(* Logix 5000 project; controller TFF vendor 1 type 14 code 107 rev 33.11; software revision 33.04; part 30 of 38 *)
(* tags used below, declared in another part *)
   Index : DINT;   // Index
   AA008 : ALIAS FOR DigitalPoint[18];
   AI101 : ALIAS FOR AnalogPoint[16];
   AI101_SIG : ALIAS FOR DigitalPoint[106];
   AI104 : ALIAS FOR AnalogPoint[17];
   AI104_SIG : ALIAS FOR DigitalPoint[107];
   AI201B : ALIAS FOR AnalogPoint[0];
   AI201B_SIG : ALIAS FOR DigitalPoint[109];
   AI202 : ALIAS FOR AnalogPoint[9];
   AI202_SIG : ALIAS FOR DigitalPoint[105];
   ARC_AI101 : ARC_pH;
   ARC_AI202 : ARC_pH;
   DF24VDC : ALIAS FOR DigitalPoint[4];
   DF24VDCPC : ALIAS FOR DigitalPoint[25];
   DF3PHP003 : ALIAS FOR DigitalPoint[27];
   DigitalInput : BOOL[256];   // Digital Input Array these bits are copied from Input cards.
   DigitalPoint : DigitalPoint[150];   // Digital Point Array
   ES001 : ALIAS FOR DigitalPoint[2];
   FI101 : ALIAS FOR AnalogPoint[19];
   FI101_SIG : ALIAS FOR DigitalPoint[110];
   MIX101 : ALIAS FOR AnalogPoint[14];
   MIX101_SIG : ALIAS FOR DigitalPoint[104];
   MIX101DF : ALIAS FOR DigitalPoint[28];
   Mixer : Mixer;   // Mixer config. structure
   Options : Options;   // Options List
   PCV101 : ALIAS FOR AnalogPoint[3];
   PCV101_SIG : ALIAS FOR DigitalPoint[102];
   PCV201 : ALIAS FOR AnalogPoint[4];
   PCV201_SIG : ALIAS FOR DigitalPoint[103];
   PI101 : ALIAS FOR AnalogPoint[6];
   PI101_SIG : ALIAS FOR DigitalPoint[98];
   PI201 : ALIAS FOR AnalogPoint[7];
   PI201_SIG : ALIAS FOR DigitalPoint[99];
   PI401 : ALIAS FOR AnalogPoint[8];
   PI401_SIG : ALIAS FOR DigitalPoint[100];
   PSH001 : ALIAS FOR DigitalPoint[21];
   PSH401 : ALIAS FOR DigitalPoint[22];
   Rack_Murr_Node0_Smart : IO_Station;   // Status of Node 0 Smart
   Rack_Murr_Node1_TFF20 : IO_Station;   // Status of Node 1 TFF20
   Rack_Murr_Node1_TFF40 : IO_Station;   // Status of Node 1 TFF40
   Rack_Murr_Node1_TFF80 : IO_Station;   // Status of Node 1 TFF80
   RSBUZZ : ALIAS FOR DigitalPoint[3];
   SIC001DF : ALIAS FOR DigitalPoint[16];
   SIC002DF : ALIAS FOR DigitalPoint[17];
   SIC003DF : ALIAS FOR DigitalPoint[29];
   TCU101 : ALIAS FOR AnalogPoint[18];
   TCU101_SIG : ALIAS FOR DigitalPoint[108];
   TCU101DF : ALIAS FOR DigitalPoint[30];
   ThisSystem : SystemType;
   TI101 : ALIAS FOR AnalogPoint[13];
   TI101_SIG : ALIAS FOR DigitalPoint[101];
   TI201 : ALIAS FOR AnalogPoint[22];
   TI201_SIG : ALIAS FOR DigitalPoint[111];
   ValveSwInput : BOOL[64];   // Valve digital input
   XS011 : ALIAS FOR DigitalPoint[14];
   XS012 : ALIAS FOR DigitalPoint[15];
   XV003 : ALIAS FOR Valve[2];
   XV004 : ALIAS FOR Valve[3];
   XV005 : ALIAS FOR Valve[4];
   XV006 : ALIAS FOR Valve[5];
   XV007 : ALIAS FOR Valve[6];
   ZS001 : ALIAS FOR DigitalPoint[6];
   ZS002 : ALIAS FOR DigitalPoint[7];
   ZS003 : ALIAS FOR DigitalPoint[8];
   ZS004 : ALIAS FOR DigitalPoint[9];
   ZS005 : ALIAS FOR DigitalPoint[10];
   ZS008 : ALIAS FOR DigitalPoint[5];
(* Process, continued *)

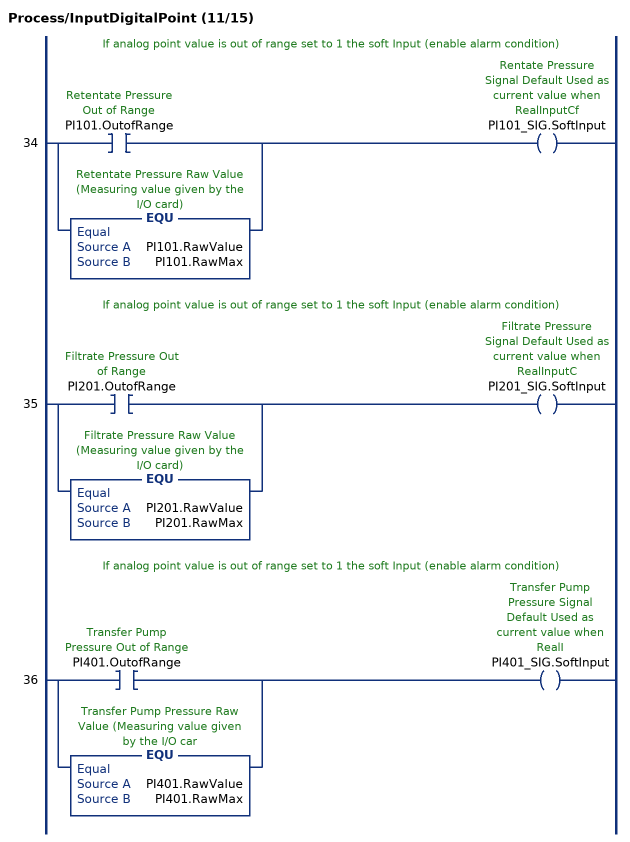
   [picture p330: Process/InputDigitalPoint rungs 34-36]
   // If analog point value is out of range set to 1 the soft Input (enable alarm condition)
   34: [XIC(PI101.OutofRange) ,EQU(PI101.RawValue,PI101.RawMax) ]OTE(PI101_SIG.SoftInput);
   // If analog point value is out of range set to 1 the soft Input (enable alarm condition)
   35: [XIC(PI201.OutofRange) ,EQU(PI201.RawValue,PI201.RawMax) ]OTE(PI201_SIG.SoftInput);
   // If analog point value is out of range set to 1 the soft Input (enable alarm condition)
   36: [XIC(PI401.OutofRange) ,EQU(PI401.RawValue,PI401.RawMax) ]OTE(PI401_SIG.SoftInput);
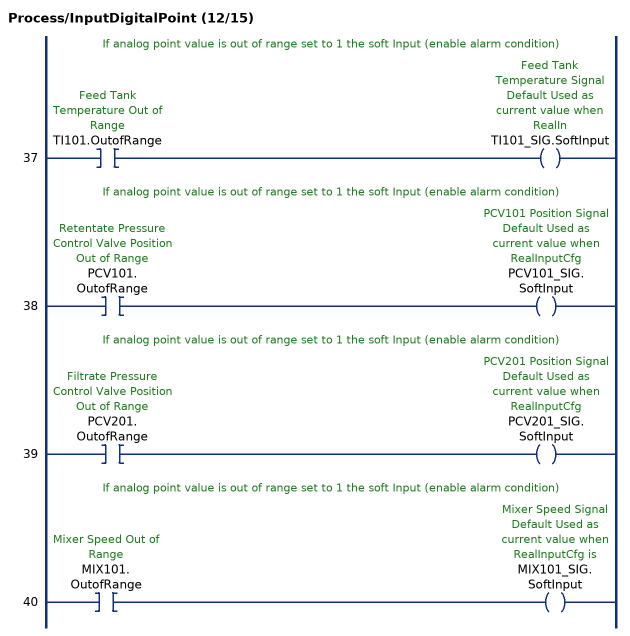
   // If analog point value is out of range set to 1 the soft Input (enable alarm condition)
   37: XIC(TI101.OutofRange)OTE(TI101_SIG.SoftInput);
   // If analog point value is out of range set to 1 the soft Input (enable alarm condition)
   38: XIC(PCV101.OutofRange)OTE(PCV101_SIG.SoftInput);
   // If analog point value is out of range set to 1 the soft Input (enable alarm condition)
   39: XIC(PCV201.OutofRange)OTE(PCV201_SIG.SoftInput);
   // If analog point value is out of range set to 1 the soft Input (enable alarm condition)
   40: XIC(MIX101.OutofRange)OTE(MIX101_SIG.SoftInput);
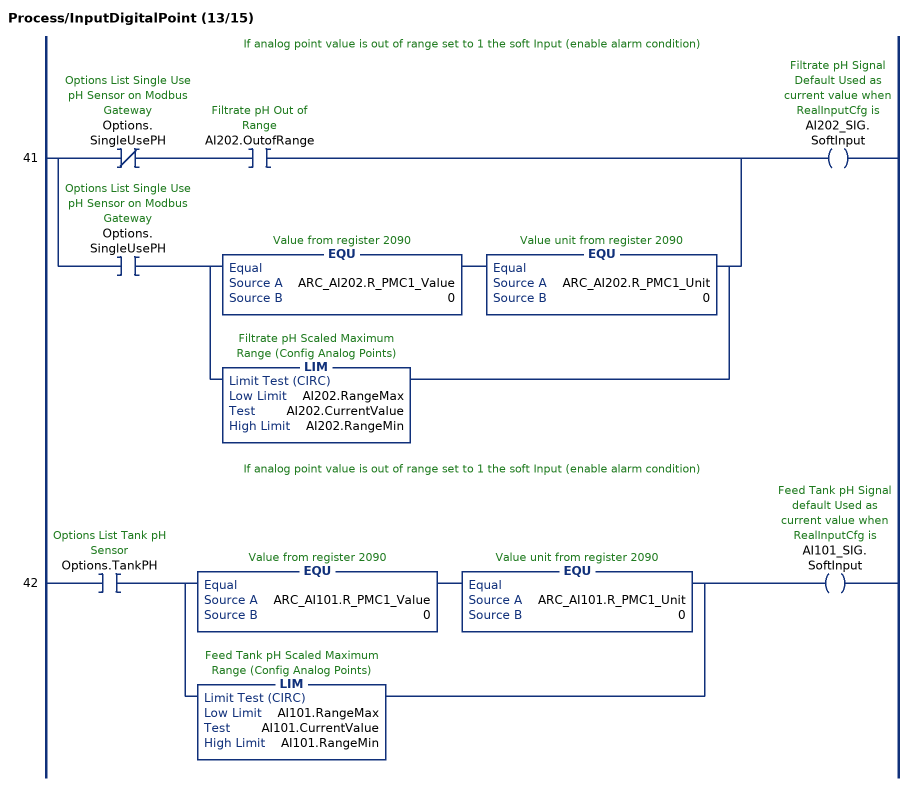
   // If analog point value is out of range set to 1 the soft Input (enable alarm condition)
   41: [XIO(Options.SingleUsePH) XIC(AI202.OutofRange) ,XIC(Options.SingleUsePH) [EQU(ARC_AI202.R_PMC1_Value,0) EQU(ARC_AI202.R_PMC1_Unit,0) ,LIM(AI202.RangeMax,AI202.CurrentValue,AI202.RangeMin) ] ]OTE(AI202_SIG.SoftInput);
   // If analog point value is out of range set to 1 the soft Input (enable alarm condition)
   42: XIC(Options.TankPH)[EQU(ARC_AI101.R_PMC1_Value,0) EQU(ARC_AI101.R_PMC1_Unit,0) ,LIM(AI101.RangeMax,AI101.CurrentValue,AI101.RangeMin) ]OTE(AI101_SIG.SoftInput);
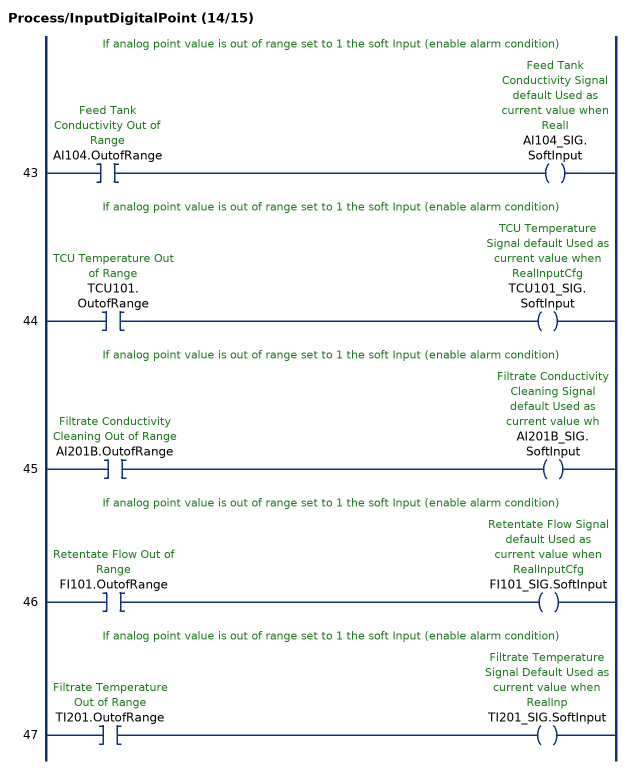
   // If analog point value is out of range set to 1 the soft Input (enable alarm condition)
   43: XIC(AI104.OutofRange)OTE(AI104_SIG.SoftInput);
   // If analog point value is out of range set to 1 the soft Input (enable alarm condition)
   44: XIC(TCU101.OutofRange)OTE(TCU101_SIG.SoftInput);
   // If analog point value is out of range set to 1 the soft Input (enable alarm condition)
   45: XIC(AI201B.OutofRange)OTE(AI201B_SIG.SoftInput);
   // If analog point value is out of range set to 1 the soft Input (enable alarm condition)
   46: XIC(FI101.OutofRange)OTE(FI101_SIG.SoftInput);
   // If analog point value is out of range set to 1 the soft Input (enable alarm condition)
   47: XIC(TI201.OutofRange)OTE(TI201_SIG.SoftInput);
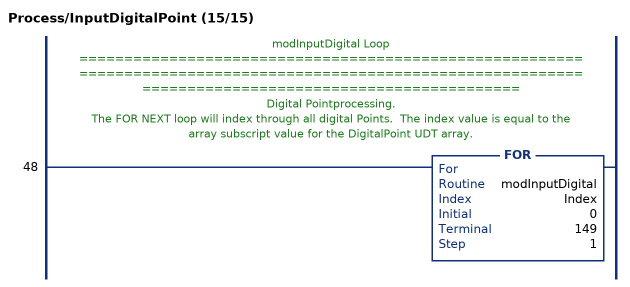
   // modInputDigital Loop
   // ==========================================================================================================================================================
   // Digital Pointprocessing.
   // The FOR NEXT loop will index through all digital Points.  The index value is equal to the array subscript value for the DigitalPoint UDT array.
   48: FOR(modInputDigital,Index,0,149,1);
END_ROUTINE

ROUTINE InputDigitalRaw   (* ladder *)
// Digital Input Routine
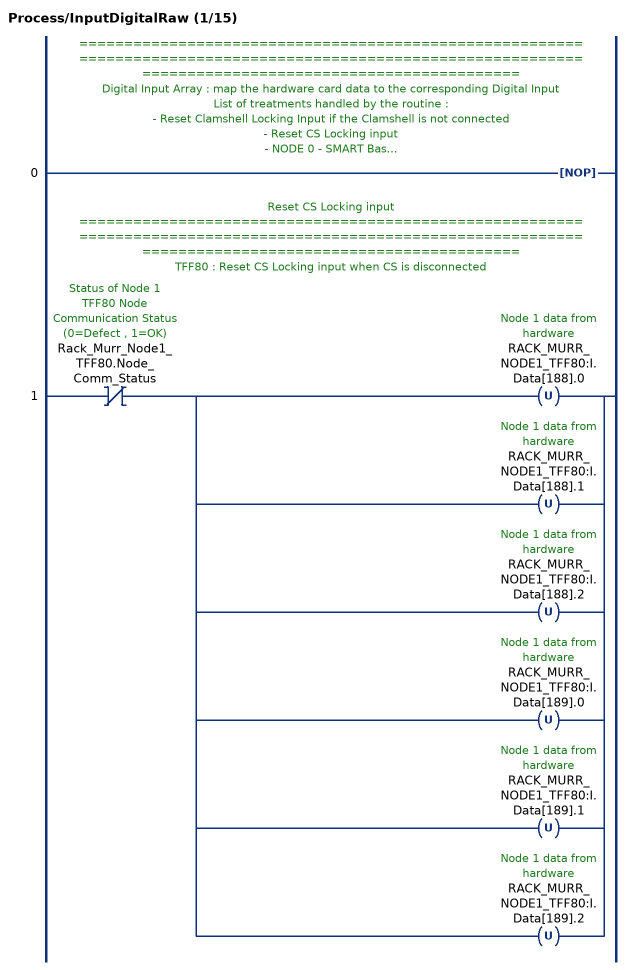
   // ==========================================================================================================================================================
   //                                                                                             Digital Input Array : map the hardware card data to the corresponding Digital Input
   //                                                     List of treatments handled by the routine :
   //                                                    - Reset Clamshell Locking Input if the Clamshell is not connected
   //                                                    - Reset CS Locking input
   //                                                    - NODE 0 - SMART Base
   //                                                         - NODE 1 - TFF80 Clamshell
   //                                                         - NODE 1 - TFF40 Clamshell
   //                                                         - NODE 1 - TFF20 Clamshell
   //                                                     -----------------------------------------------------------------------------------------------------------------------------------------------------
   //                                                     History
   // 		2019-DEC-24 - Merck - Q. Spindler - Initial version for Candidate Release 1.00.00.00.a
   // 		2020-APR-15 - Merck - Q. Spindler - Modifications for Candidate Release 1.00.00.00.b
   // - Add XS003, XS004, XS005, XS006, and XS007
   // ==========================================================================================================================================================
   0: NOP();
   // Reset CS Locking input
   // ==========================================================================================================================================================
   // TFF80 : Reset CS Locking input when CS is disconnected
   1: XIO(Rack_Murr_Node1_TFF80.Node_Comm_Status)[OTU(RACK_MURR_NODE1_TFF80:I.Data[188].0) ,OTU(RACK_MURR_NODE1_TFF80:I.Data[188].1) ,OTU(RACK_MURR_NODE1_TFF80:I.Data[188].2) ,OTU(RACK_MURR_NODE1_TFF80:I.Data[189].0) ,OTU(RACK_MURR_NODE1_TFF80:I.Data[189].1) ,OTU(RACK_MURR_NODE1_TFF80:I.Data[189].2) ];
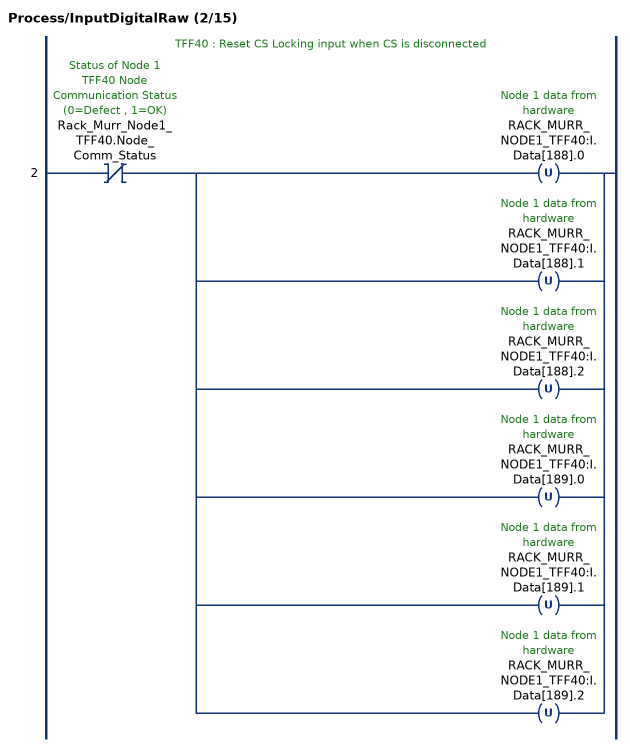
   // TFF40 : Reset CS Locking input when CS is disconnected
   2: XIO(Rack_Murr_Node1_TFF40.Node_Comm_Status)[OTU(RACK_MURR_NODE1_TFF40:I.Data[188].0) ,OTU(RACK_MURR_NODE1_TFF40:I.Data[188].1) ,OTU(RACK_MURR_NODE1_TFF40:I.Data[188].2) ,OTU(RACK_MURR_NODE1_TFF40:I.Data[189].0) ,OTU(RACK_MURR_NODE1_TFF40:I.Data[189].1) ,OTU(RACK_MURR_NODE1_TFF40:I.Data[189].2) ];
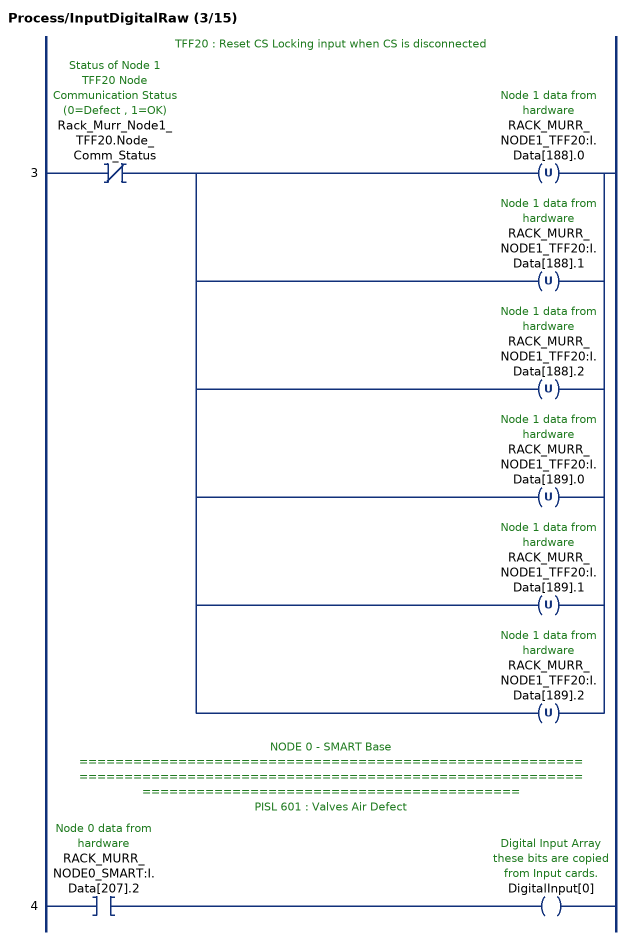
   // TFF20 : Reset CS Locking input when CS is disconnected
   3: XIO(Rack_Murr_Node1_TFF20.Node_Comm_Status)[OTU(RACK_MURR_NODE1_TFF20:I.Data[188].0) ,OTU(RACK_MURR_NODE1_TFF20:I.Data[188].1) ,OTU(RACK_MURR_NODE1_TFF20:I.Data[188].2) ,OTU(RACK_MURR_NODE1_TFF20:I.Data[189].0) ,OTU(RACK_MURR_NODE1_TFF20:I.Data[189].1) ,OTU(RACK_MURR_NODE1_TFF20:I.Data[189].2) ];
   // NODE 0 - SMART Base
   // ==========================================================================================================================================================
   // PISL 601 : Valves Air Defect
   4: XIC(RACK_MURR_NODE0_SMART:I.Data[207].2)OTE(DigitalInput[0]);
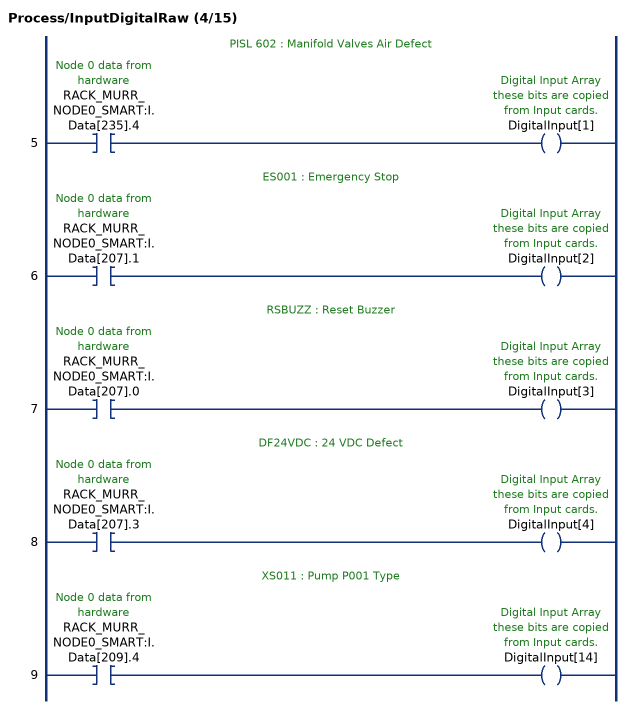
   // PISL 602 : Manifold Valves Air Defect
   5: XIC(RACK_MURR_NODE0_SMART:I.Data[235].4)OTE(DigitalInput[1]);
   // ES001 : Emergency Stop
   6: XIC(RACK_MURR_NODE0_SMART:I.Data[207].1)OTE(DigitalInput[2]);
   // RSBUZZ : Reset Buzzer
   7: XIC(RACK_MURR_NODE0_SMART:I.Data[207].0)OTE(DigitalInput[3]);
   // DF24VDC : 24 VDC Defect
   8: XIC(RACK_MURR_NODE0_SMART:I.Data[207].3)OTE(DigitalInput[4]);
   // XS011 : Pump P001 Type
   9: XIC(RACK_MURR_NODE0_SMART:I.Data[209].4)OTE(DigitalInput[14]);
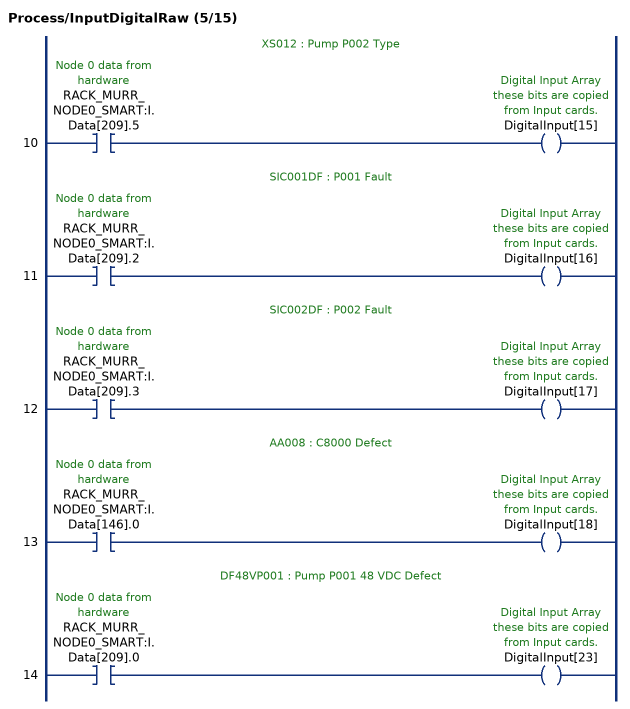
   // XS012 : Pump P002 Type
   10: XIC(RACK_MURR_NODE0_SMART:I.Data[209].5)OTE(DigitalInput[15]);
   // SIC001DF : P001 Fault
   11: XIC(RACK_MURR_NODE0_SMART:I.Data[209].2)OTE(DigitalInput[16]);
   // SIC002DF : P002 Fault
   12: XIC(RACK_MURR_NODE0_SMART:I.Data[209].3)OTE(DigitalInput[17]);
   // AA008 : C8000 Defect
   13: XIC(RACK_MURR_NODE0_SMART:I.Data[146].0)OTE(DigitalInput[18]);
   // DF48VP001 : Pump P001 48 VDC Defect
   14: XIC(RACK_MURR_NODE0_SMART:I.Data[209].0)OTE(DigitalInput[23]);
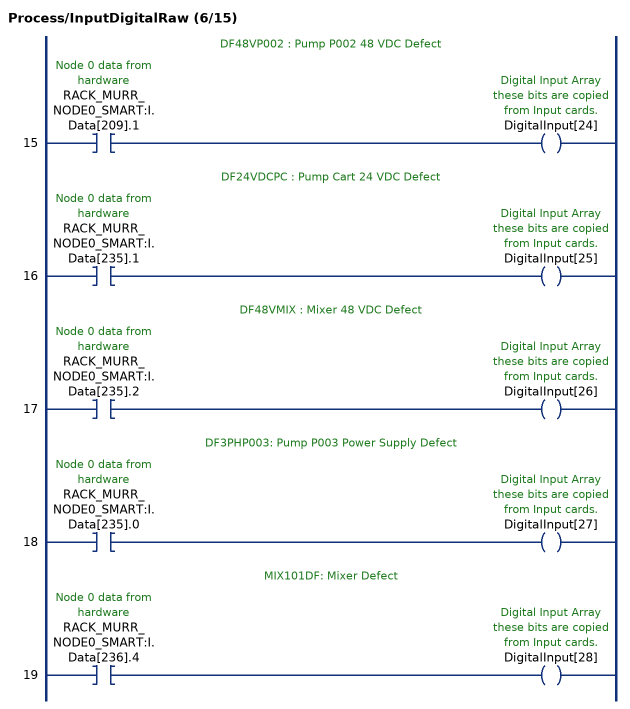
   // DF48VP002 : Pump P002 48 VDC Defect
   15: XIC(RACK_MURR_NODE0_SMART:I.Data[209].1)OTE(DigitalInput[24]);
   // DF24VDCPC : Pump Cart 24 VDC Defect
   16: XIC(RACK_MURR_NODE0_SMART:I.Data[235].1)OTE(DigitalInput[25]);
   // DF48VMIX : Mixer 48 VDC Defect
   17: XIC(RACK_MURR_NODE0_SMART:I.Data[235].2)OTE(DigitalInput[26]);
   // DF3PHP003: Pump P003 Power Supply Defect
   18: XIC(RACK_MURR_NODE0_SMART:I.Data[235].0)OTE(DigitalInput[27]);
   // MIX101DF: Mixer Defect
   19: XIC(RACK_MURR_NODE0_SMART:I.Data[236].4)OTE(DigitalInput[28]);
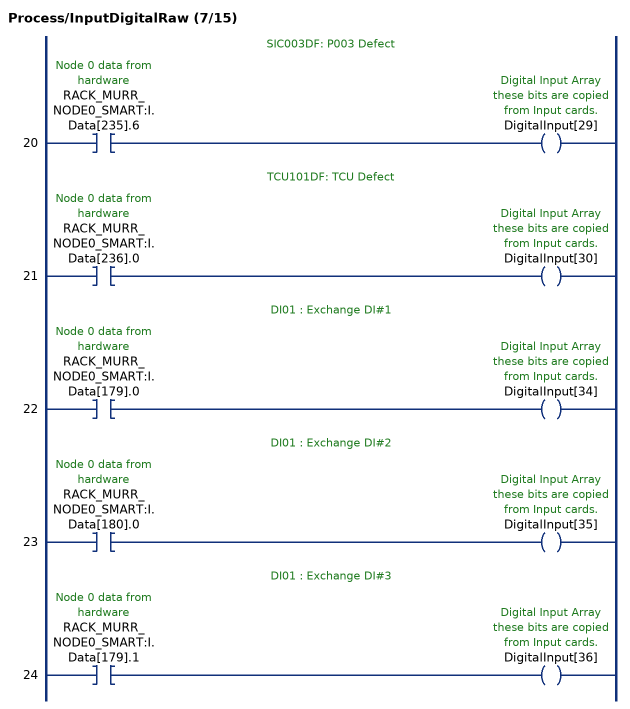
   // SIC003DF: P003 Defect
   20: XIC(RACK_MURR_NODE0_SMART:I.Data[235].6)OTE(DigitalInput[29]);
   // TCU101DF: TCU Defect
   21: XIC(RACK_MURR_NODE0_SMART:I.Data[236].0)OTE(DigitalInput[30]);
   // DI01 : Exchange DI#1
   22: XIC(RACK_MURR_NODE0_SMART:I.Data[179].0)OTE(DigitalInput[34]);
   // DI01 : Exchange DI#2
   23: XIC(RACK_MURR_NODE0_SMART:I.Data[180].0)OTE(DigitalInput[35]);
   // DI01 : Exchange DI#3
   24: XIC(RACK_MURR_NODE0_SMART:I.Data[179].1)OTE(DigitalInput[36]);
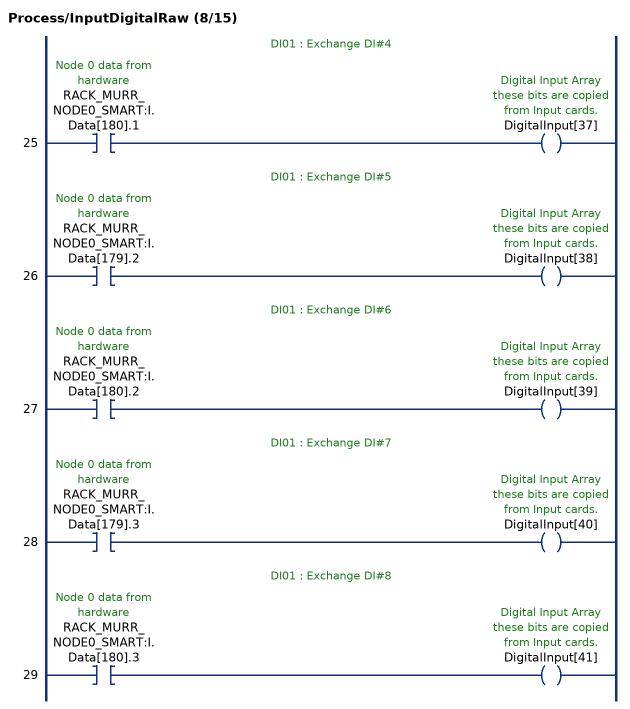
   // DI01 : Exchange DI#4
   25: XIC(RACK_MURR_NODE0_SMART:I.Data[180].1)OTE(DigitalInput[37]);
   // DI01 : Exchange DI#5
   26: XIC(RACK_MURR_NODE0_SMART:I.Data[179].2)OTE(DigitalInput[38]);
   // DI01 : Exchange DI#6
   27: XIC(RACK_MURR_NODE0_SMART:I.Data[180].2)OTE(DigitalInput[39]);
   // DI01 : Exchange DI#7
   28: XIC(RACK_MURR_NODE0_SMART:I.Data[179].3)OTE(DigitalInput[40]);
   // DI01 : Exchange DI#8
   29: XIC(RACK_MURR_NODE0_SMART:I.Data[180].3)OTE(DigitalInput[41]);
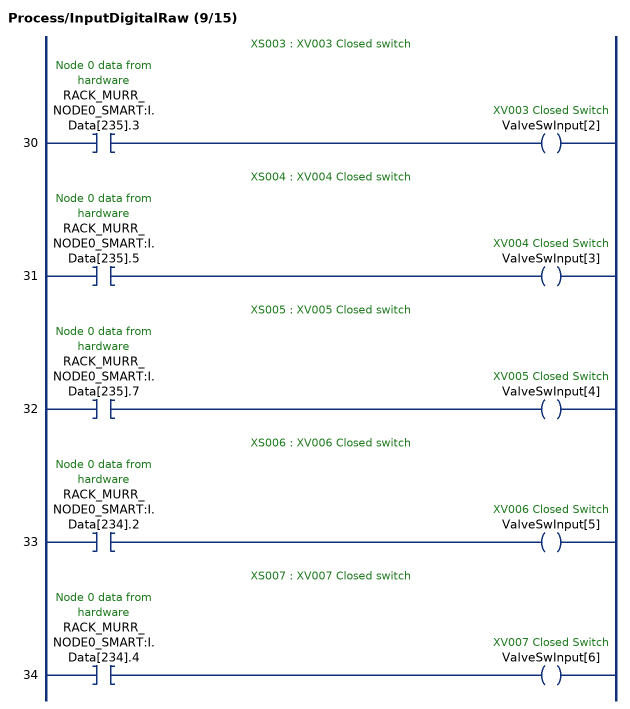
   // XS003 : XV003 Closed switch
   30: XIC(RACK_MURR_NODE0_SMART:I.Data[235].3)OTE(ValveSwInput[2]);
   // XS004 : XV004 Closed switch
   31: XIC(RACK_MURR_NODE0_SMART:I.Data[235].5)OTE(ValveSwInput[3]);
   // XS005 : XV005 Closed switch
   32: XIC(RACK_MURR_NODE0_SMART:I.Data[235].7)OTE(ValveSwInput[4]);
   // XS006 : XV006 Closed switch
   33: XIC(RACK_MURR_NODE0_SMART:I.Data[234].2)OTE(ValveSwInput[5]);
   // XS007 : XV007 Closed switch
   34: XIC(RACK_MURR_NODE0_SMART:I.Data[234].4)OTE(ValveSwInput[6]);
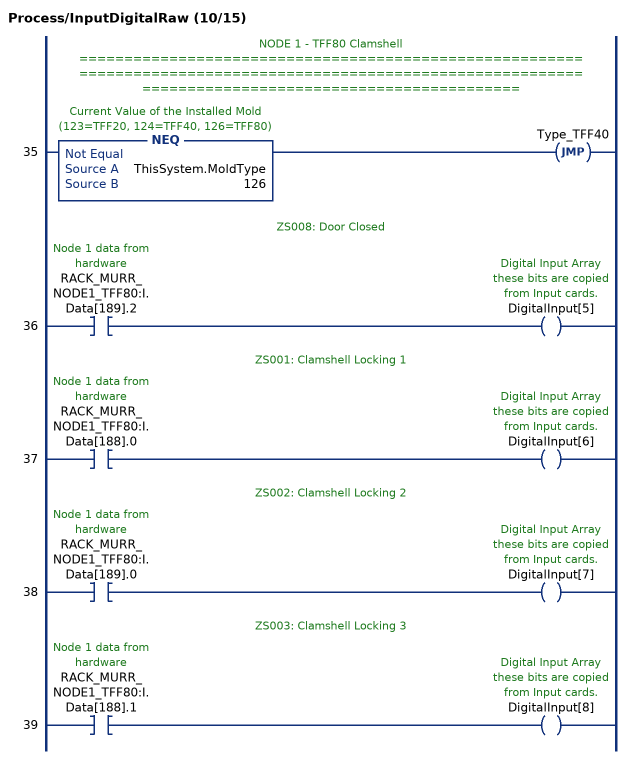
   // NODE 1 - TFF80 Clamshell
   // ==========================================================================================================================================================
   35: NEQ(ThisSystem.MoldType,126)JMP(Type_TFF40);
   // ZS008: Door Closed
   36: XIC(RACK_MURR_NODE1_TFF80:I.Data[189].2)OTE(DigitalInput[5]);
   // ZS001: Clamshell Locking 1
   37: XIC(RACK_MURR_NODE1_TFF80:I.Data[188].0)OTE(DigitalInput[6]);
   // ZS002: Clamshell Locking 2
   38: XIC(RACK_MURR_NODE1_TFF80:I.Data[189].0)OTE(DigitalInput[7]);
   // ZS003: Clamshell Locking 3
   39: XIC(RACK_MURR_NODE1_TFF80:I.Data[188].1)OTE(DigitalInput[8]);
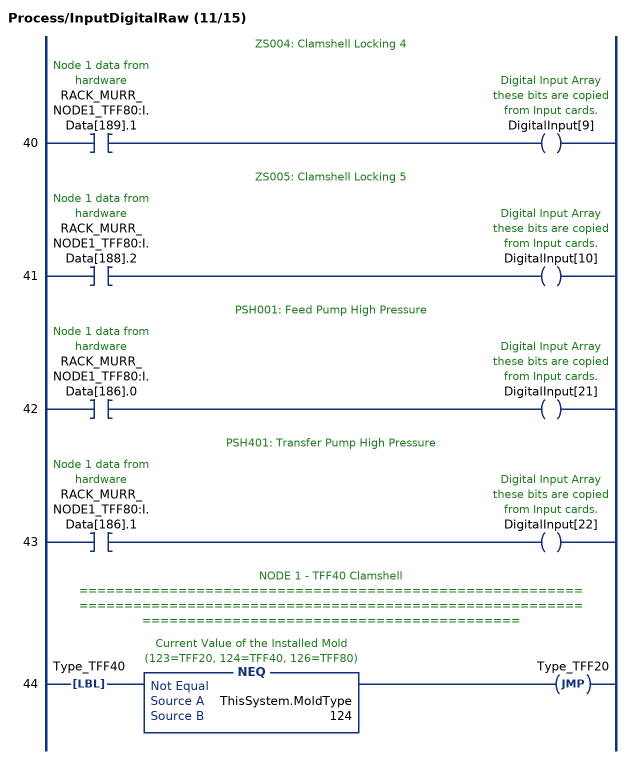
   // ZS004: Clamshell Locking 4
   40: XIC(RACK_MURR_NODE1_TFF80:I.Data[189].1)OTE(DigitalInput[9]);
   // ZS005: Clamshell Locking 5
   41: XIC(RACK_MURR_NODE1_TFF80:I.Data[188].2)OTE(DigitalInput[10]);
   // PSH001: Feed Pump High Pressure
   42: XIC(RACK_MURR_NODE1_TFF80:I.Data[186].0)OTE(DigitalInput[21]);
   // PSH401: Transfer Pump High Pressure
   43: XIC(RACK_MURR_NODE1_TFF80:I.Data[186].1)OTE(DigitalInput[22]);
   // NODE 1 - TFF40 Clamshell
   // ==========================================================================================================================================================
   44: LBL(Type_TFF40)NEQ(ThisSystem.MoldType,124)JMP(Type_TFF20);
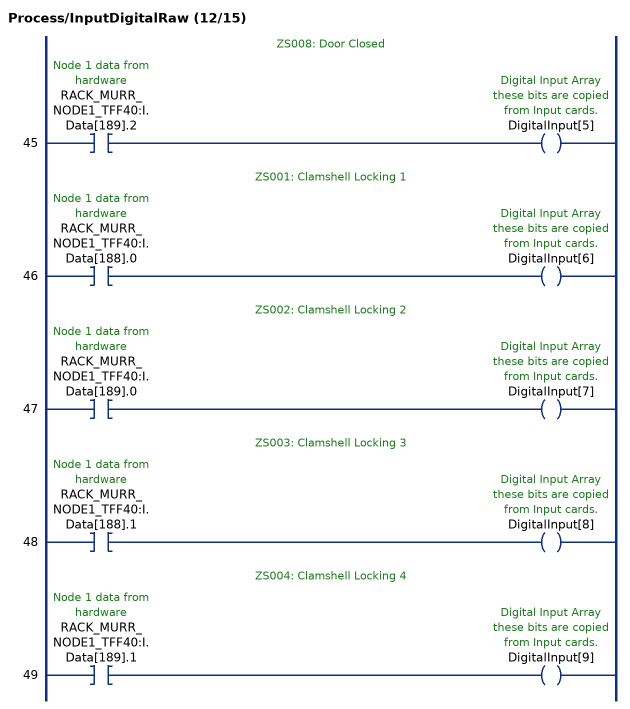
   // ZS008: Door Closed
   45: XIC(RACK_MURR_NODE1_TFF40:I.Data[189].2)OTE(DigitalInput[5]);
   // ZS001: Clamshell Locking 1
   46: XIC(RACK_MURR_NODE1_TFF40:I.Data[188].0)OTE(DigitalInput[6]);
   // ZS002: Clamshell Locking 2
   47: XIC(RACK_MURR_NODE1_TFF40:I.Data[189].0)OTE(DigitalInput[7]);
   // ZS003: Clamshell Locking 3
   48: XIC(RACK_MURR_NODE1_TFF40:I.Data[188].1)OTE(DigitalInput[8]);
   // ZS004: Clamshell Locking 4
   49: XIC(RACK_MURR_NODE1_TFF40:I.Data[189].1)OTE(DigitalInput[9]);
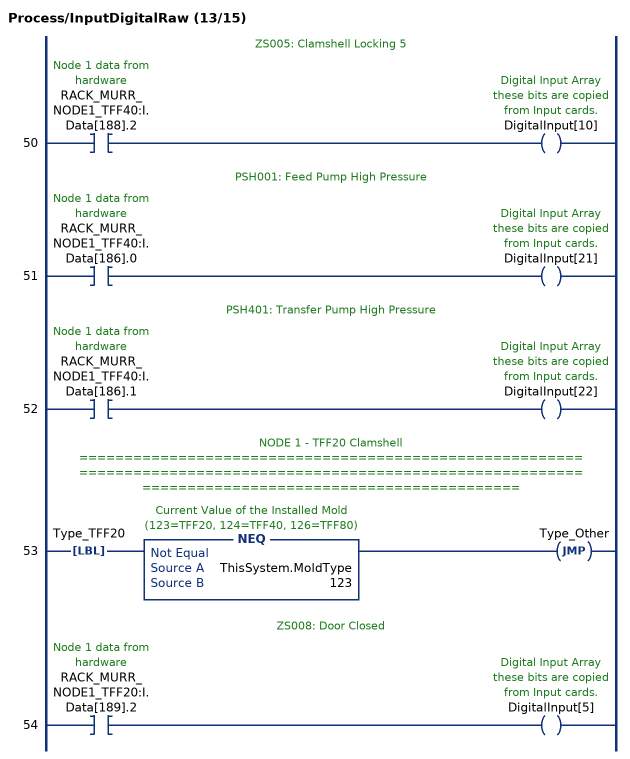
   // ZS005: Clamshell Locking 5
   50: XIC(RACK_MURR_NODE1_TFF40:I.Data[188].2)OTE(DigitalInput[10]);
   // PSH001: Feed Pump High Pressure
   51: XIC(RACK_MURR_NODE1_TFF40:I.Data[186].0)OTE(DigitalInput[21]);
   // PSH401: Transfer Pump High Pressure
   52: XIC(RACK_MURR_NODE1_TFF40:I.Data[186].1)OTE(DigitalInput[22]);
   // NODE 1 - TFF20 Clamshell
   // ==========================================================================================================================================================
   53: LBL(Type_TFF20)NEQ(ThisSystem.MoldType,123)JMP(Type_Other);
   // ZS008: Door Closed
   54: XIC(RACK_MURR_NODE1_TFF20:I.Data[189].2)OTE(DigitalInput[5]);
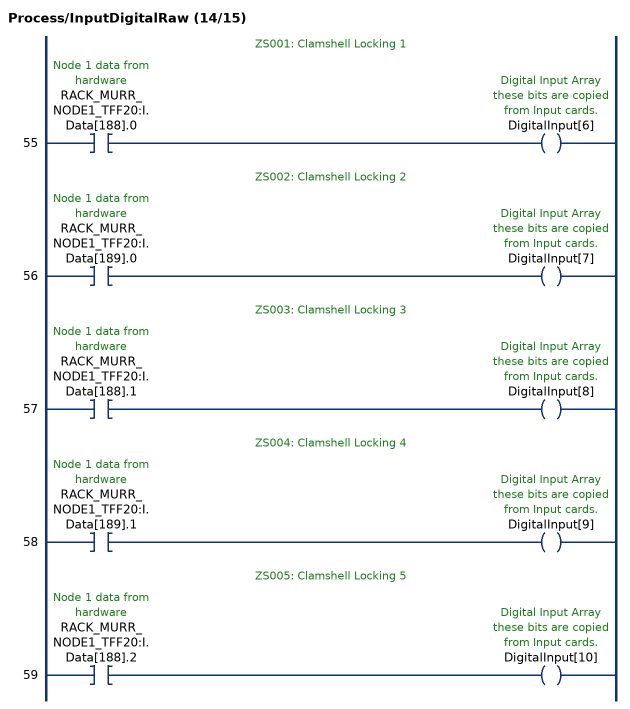
   // ZS001: Clamshell Locking 1
   55: XIC(RACK_MURR_NODE1_TFF20:I.Data[188].0)OTE(DigitalInput[6]);
   // ZS002: Clamshell Locking 2
   56: XIC(RACK_MURR_NODE1_TFF20:I.Data[189].0)OTE(DigitalInput[7]);
   // ZS003: Clamshell Locking 3
   57: XIC(RACK_MURR_NODE1_TFF20:I.Data[188].1)OTE(DigitalInput[8]);
   // ZS004: Clamshell Locking 4
   58: XIC(RACK_MURR_NODE1_TFF20:I.Data[189].1)OTE(DigitalInput[9]);
   // ZS005: Clamshell Locking 5
   59: XIC(RACK_MURR_NODE1_TFF20:I.Data[188].2)OTE(DigitalInput[10]);
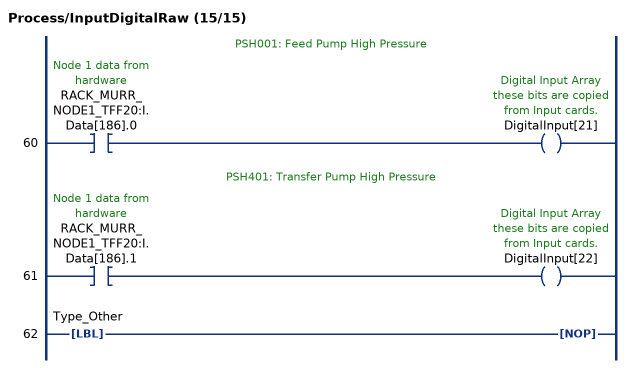
   // PSH001: Feed Pump High Pressure
   60: XIC(RACK_MURR_NODE1_TFF20:I.Data[186].0)OTE(DigitalInput[21]);
   // PSH401: Transfer Pump High Pressure
   61: XIC(RACK_MURR_NODE1_TFF20:I.Data[186].1)OTE(DigitalInput[22]);
   62: LBL(Type_Other)NOP();
END_ROUTINE
